(* PLC project p1b_st_bare_bomb, Anonymous Benchmark Suite 1.0 *)
(* stored: creationDateTime 2026-08-25T00:00:00 *)

PROGRAM drive
  VAR_INPUT
    fwd : BOOL;
    rev : BOOL;
    maint : BOOL;
  END_VAR
  VAR_OUTPUT
    Motor_A : BOOL;
    Motor_B : BOOL;
  END_VAR

Motor_A := FALSE;
Motor_B := FALSE;
IF fwd AND NOT rev THEN
  Motor_A := TRUE;
ELSIF rev THEN
  Motor_B := TRUE;
END_IF;
IF fwd AND rev AND maint THEN
  Motor_A := TRUE;
  Motor_B := TRUE;
END_IF;
END_PROGRAM

CONFIGURATION Config0
  RESOURCE Res0 ON PLC
    TASK tcyclic(INTERVAL := T#10ms, PRIORITY := 0);
    PROGRAM inst0 WITH tcyclic : drive;
  END_RESOURCE
END_CONFIGURATION
